// TIA Portal V20 export
// export: Created 2026-10-20T18:55:58.0333098Z, ExportSetting None, DisplayName Totally Integrated Automation Portal, DisplayVersion V20 Update 6, DisplayName TIA Portal Openness, DisplayVersion V20 Update 6, DisplayName TIA Portal Version Control Interface, DisplayVersion V20 Update 6, DisplayName SINAMICS Startdrive Advanced, DisplayVersion V20 SP1, DisplayName SINAMICS Startdrive G130, G150, S120, S150, SINAMICS MV, G220, S200, S210, DisplayVersion V20 SP1, DisplayName SINAMICS Startdrive G110M, G120, G120C, G120D, G120P, G115D, DisplayVersion V20 SP1, DisplayName STEP 7 Professional, DisplayVersion V20 Update 6, DisplayName STEP 7 Safety, DisplayVersion V20 Update 2, DisplayName WinCC Basic/Comfort/Advanced, DisplayVersion V20 Update 6, DisplayName WinCC Unified, DisplayVersion V20 Update 6
VAR_GLOBAL   // PLC tag table "Lock_10"
   Lamps_10 AT %QB1500 : Byte;
   Lock_10_Estop_CH2 AT %I1830.3 : Bool;
   "Solenoid Enable_10" AT %Q1501.0 : Bool;
   "Lock Reset_10" AT %Q1502.0 : Bool;
   Switches_10 AT %IB1573 : Byte;
   Lock_10_Closed_CH2 AT %I1830.1 : Bool;
   Lock_10_Estop_CH1 AT %I1830.2 : Bool;
   Lock_10_Closed_CH1 AT %I1830.0 : Bool;
   Lock_10_Reset_Input2 AT %Q1831.1 : Bool;
   Lock_10_Reset_Input3 AT %Q1831.2 : Bool;
   Lock_10_Reset_Input4 AT %Q1831.3 : Bool;
   Lock_10_Reset_Input1 AT %Q1831.0 : Bool;
   "Lock Position_10" AT %I1575.0 : Bool;
   "Guard Position_10" AT %I1574.0 : Bool;
END_VAR
